{attribute 'no_assign'}
FUNCTION_BLOCK FB_WTURBINEServerSession IMPLEMENTS I_ScsmAbortIndEventSink, I_ScsmAssociateIndEventSink, I_ScsmReleaseIndEventSink
VAR_INPUT
	fbConnection		: FB_iec61850ConnectionClass := (ipAbortInd:=THIS^, ipAssociateInd:=THIS^, ipReleaseInd:=THIS^);
	nID					: UDINT;
END_VAR
VAR
	_bAbort				: BOOL; (* Rising edge activates AbortReq() command execution *)
	_bDisconnect		: BOOL; (* Rising edge activates ReleaseReq() command execution *)
	
	state				: BYTE;
	eState				: E_AsyncEnvironmentState; (* Environment state *)
	eLinkStatus			: E_ScsmLinkStatus; (* Network adapter link status *)
	bBusy				: BOOL; (* If TRUE => command execution is busy *)
	bSuccess			: BOOL;
	ipResult			: I_AsyncServiceResultClass;
	sLastErrorResult	: T_MaxString;
	fbAbortReason		: FB_ServiceErrorClass := (stError:=SUCCESS_EVENT);
	sLastAbortReason	: T_MaxString;
END_VAR

fbConnection.Execute();
eState:= fbConnection.eState;
eLinkStatus:= fbConnection.eLinkStatus;

(* Execute control model control block implementations *)
// fbWTURBINE.WTURBINELD0.LLN0.Mod_.fbControl.Execute();
// fbWTURBINE.WTURBINELD0.WTUR1.CmdBlk.fbControl.Execute();
// fbWTURBINE.WTURBINELD0.WNAC1.CtlMd.fbControl.Execute();
// fbWTURBINE.WTURBINELD0.WYAW1.YwBrk.fbControl.Execute();

// fbWTURBINE[nID].WTURBINELD0.LLN0.Mod_.fbControl.Execute();
// fbWTURBINE[nID].WTURBINELD0.WTUR1.CmdBlk.fbControl.Execute();
// fbWTURBINE[nID].WTURBINELD0.WNAC1.CtlMd.fbControl.Execute();
// fbWTURBINE[nID].WTURBINELD0.WYAW1.YwBrk.fbControl.Execute();
// fbWTURBINE[nID].WTURBINELD0.WTUR1.DmdWSpt.fbControl.Execute();

(* Execute server control block implementations *)
fbWTURBINE[nID].WTURBINELD0.WPPD1.urcb01.Server.Execute();

fbWTURBINE[nID].WTURBINELD0.LLN0.Mod_.fbControl.Execute();
fbWTURBINE[nID].WTURBINELD0.WTUR1.TurOp.st_.fbControl.Execute();
fbWTURBINE[nID].WTURBINELD0.WTUR1.TurCtl.st_.fbControl.Execute();
fbWTURBINE[nID].WTURBINELD0.WTUR1.DmdWSpt.val.fbControl.Execute();
fbWTURBINE[nID].WTURBINELD0.WYAW1.YwAngSpt.val.fbControl.Execute();
fbWTURBINE[nID].WTURBINELD0.WPPD1.DevOp.st_.fbControl.Execute();
fbWTURBINE[nID].WTURBINELD0.WPPD1.ClrOp.st_.fbControl.Execute();

CASE state OF
	0: (* Initial state *)
		IF _bAbort THEN (* Abort connection => execute AbortReq() command *)
			_bAbort:= FALSE;
			bSuccess:= fbConnection.AbortReq(ipReason:=fbAbortReason, ipSink:=0, ipResult=>ipResult);
			state:= SEL(bSuccess, 100, 1);
		ELSIF eState = E_AsyncEnvironmentState.Established AND _bDisconnect THEN (* Close/release connection => execute ReleaseReq() command *)
			_bDisconnect:= FALSE;
			bSuccess:= fbConnection.ReleaseReq(ipSink:=0, ipResult=>ipResult);
			state:= SEL(bSuccess, 100, 1);
		ELSIF eState = E_AsyncEnvironmentState.Established THEN (* Connection established => exchange IED data *)
			state:= 10;
		END_IF
		_bDisconnect:= FALSE;
		(*==================================================================================================================================================================*)
	1: (* Wait for AbortReq() or ReleaseReq() command completion *)
		IF ipResult <> 0 THEN
			ipResult.Execute();
			IF NOT (bBusy:=ipResult.IsBusy()) THEN
				state:= SEL(ipResult.IsCompleted(), 100(* failed or aborted *), 0(* succeeded *));
			END_IF
		END_IF
		(*==================================================================================================================================================================*)
	10: (* connection established *)
		state:= 0;
		(*==================================================================================================================================================================*)
	100: (* Error state *)
		state:= 0;
		IF ipResult <> 0 THEN
			sLastErrorResult:= ipResult.Dump();
		END_IF
END_CASE

PROPERTY bAbort : BOOL
SET
_bAbort:= bAbort;
END_SET
END_PROPERTY

PROPERTY bDisconnect : BOOL
SET
_bDisconnect:= bDisconnect;
END_SET
END_PROPERTY

(* This method receives IEC61850::Abort.ind primitive. *)
METHOD OnAbortInd
VAR_INPUT
	ipAA		: I_ScsmAssociationClass; (* Application association. If = 0 => optional. *)
	bPAbort		: BOOL; (* TRUE => P-Abort.request(), issued by provider, FALSE => Abort.request(), issued by user. *)
	ipReason	: I_ServiceErrorClass; (* Abort reason. *)
	ipData		: I_BaseStreamClass; (* Optional data. If = 0 => default, no data. *)
END_VAR
VAR
END_VAR
IF ipReason <> 0 THEN
	sLastAbortReason:= ipReason.Dump();
END_IF
END_METHOD

(* This method receives IEC61850::Associate.ind primitive. *)
METHOD OnAssociateInd : BOOL
VAR_INPUT
	ipAA			: I_ScsmAssociationClass; (* Application association. If = 0 => optional. *)
END_VAR
VAR_OUTPUT
	ipResult		: I_AsyncServiceResultClass; (* Interface pointer to service state and result information *)
END_VAR
VAR
END_VAR
sLastAbortReason:= '';
sLastErrorResult:= '';
OnAssociateInd:= fbConnection.AssociateRsp(ipResult=>ipResult);
END_METHOD

(* This method receives IEC61850::Release.ind primitive. *)
METHOD OnReleaseInd : BOOL
VAR_INPUT
	ipAA	: I_ScsmAssociationClass; (* Application association. If = 0 => optional. *)
END_VAR
VAR_OUTPUT
	ipResult: I_AsyncServiceResultClass;
END_VAR
VAR
END_VAR
OnReleaseInd:= fbConnection.ReleaseRsp(ipResult=>ipResult);
END_METHOD

END_FUNCTION_BLOCK

(* stored: Version 1.1.0.1
   POU FB_WTURBINEServerSession: Id {52982ed7-c084-408a-b17e-4762296c4a91}, SpecialFunc None
   Property bAbort: Id {97d8b437-d2c9-47cd-82ea-a6b954c980d6}
   Set Set: Id {ca5258cf-1c1a-4767-8103-8f21380a60dd}
   Property bDisconnect: Id {9c1ed6a7-54ab-4759-9332-5c6b35762260}
   Set Set: Id {d6828e8d-2e85-4d8d-995d-35d55ff15c90}
   Method OnAbortInd: Id {3f571836-fd18-4535-a54e-fd567c3a0ce9}
   Method OnAssociateInd: Id {5129c690-b655-4fbc-b37f-d6f0501f092f}
   Method OnReleaseInd: Id {f690f31c-8611-4010-8e94-ea002193ebee} *)
